FUNCTION_BLOCK logiBUS_QD_FREQ (* Output service interface function block for a frequency output (MCPWM, duty cycle 50 %, frequency in mHz in DWORD) *)
  (* Standard: 61499-2; Description: Copyright (c) 2026 HR Agrartechnik GmbH This program and the accompanying materials are made available under the terms of the Eclipse Public License 2.0 which is available at https://www.eclipse.org/legal/epl-2.0/ SPDX-License-Identifier: EPL-2.0 *)
  (* Version 1.0, 2026-11-06, Franz Höpfinger, HR Agrartechnik GmbH, initial version *)
  PACKAGE logiBUS::io::DQ;
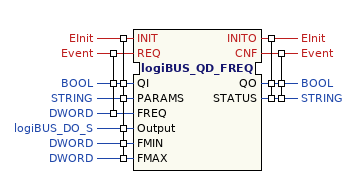
  EVENT_INPUT
    INIT : EInit WITH QI, PARAMS, Output, FMIN, FMAX; (* Service Initialization *)
    REQ WITH QI, FREQ; (* Service Request *)
  END_EVENT
  EVENT_OUTPUT
    INITO : EInit WITH QO, STATUS; (* Initialization Confirm *)
    CNF WITH QO, STATUS; (* Confirmation of Requested Service *)
  END_EVENT
  VAR_INPUT
    QI : BOOL; (* Event Input Qualifier *)
    PARAMS : STRING; (* Service Parameters *)
    FREQ : DWORD; (* Frequency in mHz (1000 = 1 Hz) like ISOBUS DDI 583 Setpoint Frequency (resolution 0.001 Hz). 0 = output off (low). Duty cycle fixed 50 %. Values outside FMIN..FMAX are limited, STATUS says so. Takes effect at the end of the running period (no glitch). Power stage limits, not checked: APIXON 15 PWR Q1 (BTH50030) max. 100 Hz; BTS7030/BTT6030/BTH6070 some 100 Hz; Trainer20 without power stage *)
    Output : logiBUS::io::DQ::logiBUS_DO_S := logiBUS_DO::Invalid; (* Identify the Output Output_Q1..Q8 *)
    FMIN : DWORD := 10000; (* Lowest frequency in mHz, read at INIT. Sets the timer resolution (16-bit timer: resolution = about FMIN * 65536): the higher FREQ is above FMIN, the coarser the steps (step about FREQ^2 / resolution). Default 10 Hz: 640 kHz resolution, step 1.6 Hz at 1 kHz, 156 Hz at 10 kHz *)
    FMAX : DWORD := 10000000; (* Highest frequency in mHz, read at INIT. FREQ above it is limited. Never more than the chip can produce with the resolution from FMIN (half the resolution) *)
  END_VAR
  VAR_OUTPUT
    QO : BOOL; (* Event Output Qualifier *)
    STATUS : STRING; (* Service Status *)
  END_VAR
END_FUNCTION_BLOCK
